TYPE ST_Tank_Level :
STRUCT
	//Input signals fro I/O
	bIn_LL_signal	:	BOOL :=TRUE	;
	bIn_HL_signal	:	BOOL :=TRUE	;
	//Tank level state, empty, Low level, High level
	e_state			:	E_Tank_Level:=E_Tank_Level.eHL	;
	
	rTankLevel				:	REAL	;
	rTankLevelPercentage	:	REAL	;
END_STRUCT
END_TYPE

(* stored: Version 1.1.0.1, ProductVersion 3.1.4024.12
   DUT ST_Tank_Level: Id {64e2480b-23b8-45ca-9775-ddf4648b5222} *)
